Fanuc KAREL source: KT00724.KL

PROGRAM KT00724
%NOLOCKGROUP
VAR
  P1: JOINTPOS
  P2: JOINTPOS
  OUT: BOOLEAN
BEGIN
  OUT = UNINIT(P1)
END KT00724
